Fanuc KAREL source: kb00045.KL

PROGRAM KB00045
%STACKSIZE=65535
%PRIORITY=65535
%NOLOCKGROUP
VAR
P1 : STRING[80]
P2 : INTEGER
BEGIN
P1='A'
P2=1
CONT_TASK(P1,P2)
END KB00045
